// TIA Portal V20 export
// export: Created 2026-10-19T18:36:07.770405Z, ExportSetting WithDefaults, DisplayName Totally Integrated Automation Portal, DisplayVersion V20 Update 6, DisplayName TIA Portal Openness, DisplayVersion V20 Update 6, DisplayName TIA Portal Version Control Interface, DisplayVersion V20 Update 6, DisplayName SINAMICS Startdrive Advanced, DisplayVersion V20 SP1, DisplayName SINAMICS Startdrive G130, G150, S120, S150, SINAMICS MV, G220, S200, S210, DisplayVersion V20 SP1, DisplayName SINAMICS Startdrive G110M, G120, G120C, G120D, G120P, G115D, DisplayVersion V20 SP1, DisplayName STEP 7 Professional, DisplayVersion V20 Update 6, DisplayName STEP 7 Safety, DisplayVersion V20 Update 2, DisplayName WinCC Basic/Comfort/Advanced, DisplayVersion V20 Update 6, DisplayName WinCC Unified, DisplayVersion V20 Update 6
FUNCTION "Feed_Steptable_FC" : Void   // FC44, SCL
{ S7_Optimized_Access := 'TRUE' }
VERSION : 0.1
// stored: AutoNumber true, IsIECCheckEnabled false, SetENOAutomatically false, UDAEnableTagReadback false
   VAR_INPUT
      CurrentTime : String;
      Task_Type : Int;
      Source_Location : DInt;
      Destination_Location : DInt;
      Shuttle_ID : Int;
   END_VAR
   VAR_IN_OUT
      StepTable : "OrderTable_UDT";
   END_VAR
BEGIN
   #StepTable.OrderNo := "OrderNo" + 1;
   #StepTable.StepNo := "OrderNo" + 1;
   #StepTable.PlaceTime := #CurrentTime;

   #StepTable.OPC_Control.Task_ID := "OrderNo" + 1;
   #StepTable.OPC_Control.Task_Type := #Task_Type;
   #StepTable.OPC_Control.Source_Location := #Source_Location;
   #StepTable.OPC_Control.Destination_Location := #Destination_Location;
   #StepTable.OPC_Control.Shuttle_ID := #Shuttle_ID;
END_FUNCTION
